Fanuc KAREL source: kt00710.KL

PROGRAM KT00710
%STACKSIZE=65535
%PRIORITY=65535
%NOLOCKGROUP
VAR
B1 : BOOLEAN
B2 : BOOLEAN
OUT : BOOLEAN
BEGIN
B1=TRUE
B2=FALSE
B1=TRUE
B2=FALSE
-- UNRESOLVED_PC line 12 opcodes [22 63 23] marker_code=48
END KT00710
